{attribute 'Tc2GvlVarNames'}
VAR_GLOBAL
	stgGr00HMI			:ST_Gr00HMIRef;
END_VAR

(* stored: Version 1.1.0.1, ProductVersion 3.1.4024.15
   GVL GVL_Gr00HMI: Id {98092ee8-3520-4779-a50e-0065a8257650} *)
